FUNCTION_BLOCK FsDir (* List a directory of the file server *)
  (* Standard: 61499-2; Description: Uses iso_FscOpenFile() (directory), iso_FscReadFile() and iso_FscCloseFile() of the CCI ISOBUS driver (ISO 11783-13). \n The smallest of the four arrays is the limit. More entries give ERR with s16Status E_OVERFLOW; the arrays then hold the first entries. \n adtModified is the local time of the server as stored on the medium (FAT, 2 s). \n Client is NmDestin.s16OwnCfHnd, file server is NmDestin.s16Handle (e.g. found with NmGetCfInfo, NAME function 61). \n The FB opens its own io channel to the server and closes it at the end. One job at a time: REQ during a job gives ERR with s16Status E_BUSY. \n Every REQ ends with exactly one CNF or ERR. *)
  (* Version 1.0, 2026-11-26, Franz Höpfinger, initial API and implementation and/or initial documentation *)
  PACKAGE isobus::fs;
  IMPORT isobus::pgn::ISONETEVENT_T;
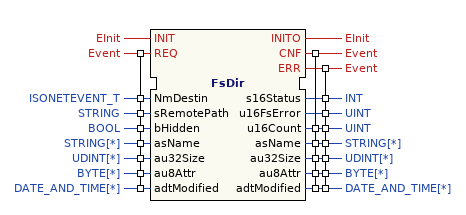
  EVENT_INPUT
    INIT : EInit; (* Service Initialization *)
    REQ WITH NmDestin, sRemotePath, bHidden, asName, au32Size, au8Attr, adtModified; (* List the directory *)
  END_EVENT
  EVENT_OUTPUT
    INITO : EInit; (* Initialization Confirm *)
    CNF WITH u16Count, asName, au32Size, au8Attr, adtModified; (* Directory listed *)
    ERR WITH s16Status, u16FsError, u16Count, asName, au32Size, au8Attr, adtModified; (* Job failed *)
  END_EVENT
  VAR_INPUT
    NmDestin : isobus::pgn::ISONETEVENT_T; (* Client (s16OwnCfHnd) and file server (s16Handle) *)
    sRemotePath : STRING; (* Directory on the file server, e.g. data or \\USB\ *)
    bHidden : BOOL; (* TRUE: list hidden entries too *)
  END_VAR
  VAR_OUTPUT
    s16Status : INT; (* With ERR: driver return value or own error (E_BUSY, E_RANGE, E_CONFIG) *)
    u16FsError : UINT; (* With ERR: file server or client error (ISO 11783-13 B.9, 6400 ff. client) *)
    u16Count : UINT; (* Number of entries in the arrays *)
  END_VAR
  VAR_IN_OUT
    asName : ARRAY [*] OF STRING; (* Names *)
    au32Size : ARRAY [*] OF UDINT; (* Sizes in bytes *)
    au8Attr : ARRAY [*] OF BYTE; (* Attributes: 16#10 directory, 16#01 read-only, 16#02 hidden *)
    adtModified : ARRAY [*] OF DATE_AND_TIME; (* Last change *)
  END_VAR
END_FUNCTION_BLOCK
